Staubli VAL3: fermerPince.pgx

program fermerPince()
begin
  open(tPince)
end
